Fanuc KAREL source: KT00656.KL

PROGRAM KT00656
%NOLOCKGROUP
VAR
  P1: POSITION
  P2: POSITION
  OUT: REAL
BEGIN
  OUT = + P1
END KT00656
